// TIA Portal V21 export
TagTable "Pump"
  PumpSpeed : Int  (%MW10, @Connection@, 1 s)
  PumpOn : Bool  (%M0.0, @Connection@, 100 ms)
  Flow : Real  (%MD20, @Connection@, 500 ms)
  SpeedSetpoint : Int  ()
